FUNCTION_BLOCK FB_EL3312ChannelDiagnosis_1
VAR_INPUT
	stChannelState				:ST_EL3312ChannelState;
END_VAR
VAR_OUTPUT
	bChannelOK					:BOOL;
	bLimit1						:BOOL;			(* State limit 1 *)
	bLimit2 						:BOOL;			(* State limit 2 *)
END_VAR
VAR

END_VAR


(* General Channel Status *)
IF stChannelState.bUnderrange = 0
    AND stChannelState.bOverrange = 0
    AND stChannelState.bError = 0
    AND stChannelState.bState = 0
THEN
	bChannelOK := TRUE;
ELSE
	bChannelOK := FALSE;
END_IF

(*bLimit1 := stChannelState.byLimit1;
bLimit2 := stChannelState.byLimit2*);

END_FUNCTION_BLOCK

(* stored: Version 1.1.0.1, ProductVersion 3.1.4024.15
   POU FB_EL3312ChannelDiagnosis_1: Id {81d5856e-dc34-4356-8cdb-3f3d78c0192d}, SpecialFunc None *)
